TYPE stLightColor :
STRUCT
	Red : USINT;
	Green : USINT;
	Blue : USINT;
END_STRUCT
END_TYPE

(* stored: Version 1.1.0.1
   DUT stLightColor: Id {bfd7d273-8fc8-4cff-b04a-2c525a61ab96} *)
